TYPE "DT_PAR_PID_CROSS_FLOW_VALVE_1"
VERSION : 0.1
   STRUCT
      INPUT_RAMP_MIN_VAL { S7_SetPoint := 'False'} : "DT_PARAM_SOLO" := (FALSE, 832, 0, 0.0, 0, T#0MS, 0.0, 0.0, '%');
      INPUT_RAMP_MAX_VAL { S7_SetPoint := 'False'} : "DT_PARAM_SOLO" := (FALSE, 833, 0, 0.0, 0, T#0MS, 0.0, 0.0, '%');
      INPUT_RAMP_FALLING_TIME { S7_SetPoint := 'False'} : "DT_PARAM_SOLO" := (FALSE, 834, 0, 0.0, 0, T#0MS, 0.0, 0.0, 's');
      INPUT_RAMP_RISING_TIME { S7_SetPoint := 'False'} : "DT_PARAM_SOLO" := (FALSE, 835, 0, 0.0, 0, T#0MS, 0.0, 0.0, 's');
      OUTPUT_RAMP_FALLING_TIME { S7_SetPoint := 'False'} : "DT_PARAM_SOLO" := (FALSE, 836, 0, 0.0, 0, T#0MS, 0.0, 0.0, 's');
      OUTPUT_RAMP_RISING_TIME { S7_SetPoint := 'False'} : "DT_PARAM_SOLO" := (FALSE, 837, 0, 0.0, 0, T#0MS, 0.0, 0.0, 's');
      MAN_ON { S7_SetPoint := 'False'} : "DT_PARAM_SOLO" := (FALSE, 838, 1, 0.0, 0, T#0MS, 0.0, 0.0, '-');
      P_SEL { S7_SetPoint := 'False'} : "DT_PARAM_SOLO" := (FALSE, 839, 1, 0.0, 0, T#0MS, 0.0, 0.0, '-');
      I_SEL { S7_SetPoint := 'False'} : "DT_PARAM_SOLO" := (FALSE, 840, 1, 0.0, 0, T#0MS, 0.0, 0.0, '-');
      INT_HOLD { S7_SetPoint := 'False'} : "DT_PARAM_SOLO" := (FALSE, 841, 1, 0.0, 0, T#0MS, 0.0, 0.0, '-');
      D_SEL { S7_SetPoint := 'False'} : "DT_PARAM_SOLO" := (FALSE, 842, 1, 0.0, 0, T#0MS, 0.0, 0.0, '-');
      NUM_OF_CYCLES { S7_SetPoint := 'False'} : "DT_PARAM_SOLO" := (FALSE, 843, 1, 0.0, 0, T#0MS, 0.0, 0.0, '-');
      GAIN { S7_SetPoint := 'False'} : "DT_PARAM_SOLO" := (FALSE, 844, 0, 0.0, 0, T#0MS, 0.0, 0.0, '');
      TI { S7_SetPoint := 'False'} : "DT_PARAM_SOLO" := (FALSE, 845, 1, 0.0, 0, T#0MS, 0.0, 0.0, '-');
      TD { S7_SetPoint := 'False'} : "DT_PARAM_SOLO" := (FALSE, 846, 1, 0.0, 0, T#0MS, 0.0, 0.0, '-');
      TM_LAG { S7_SetPoint := 'False'} : "DT_PARAM_SOLO" := (FALSE, 847, 1, 300.0, 0, T#0MS, 0.0, 0.0, '-');
      DEAD_W { S7_SetPoint := 'False'} : "DT_PARAM_SOLO" := (FALSE, 848, 0, 100.0, 0, T#0MS, 0.0, 0.0, '%');
      LMN_HLM { S7_SetPoint := 'False'} : "DT_PARAM_SOLO" := (FALSE, 849, 0, 30.0, 0, T#0MS, 0.0, 0.0, '%');
      LMN_LLM { S7_SetPoint := 'False'} : "DT_PARAM_SOLO" := (FALSE, 850, 0, 300.0, 0, T#0MS, 0.0, 0.0, '%');
      REF_MIN_VAL { S7_SetPoint := 'False'} : "DT_PARAM_SOLO" := (FALSE, 851, 0, 0.0, 0, T#0MS, 0.0, 0.0, '%');
      REF_MAX_VAL { S7_SetPoint := 'False'} : "DT_PARAM_SOLO" := (FALSE, 852, 0, 0.0, 0, T#0MS, 0.0, 0.0, '%');
      LMN_FAC { S7_SetPoint := 'False'} : "DT_PARAM_SOLO" := (FALSE, 853, 0, 0.0, 0, T#0MS, 0.0, 0.0, '-');
      LMN_OFFSET { S7_SetPoint := 'False'} : "DT_PARAM_SOLO" := (FALSE, 854, 0, 0.0, 0, T#0MS, 0.0, 0.0, '%');
      DISV { S7_SetPoint := 'False'} : "DT_PARAM_SOLO" := (FALSE, 855, 0, 0.0, 0, T#0MS, 0.0, 0.0, '-');
      MAN { S7_SetPoint := 'False'} : "DT_PARAM_SOLO" := (FALSE, 856, 0, 0.0, 0, T#0MS, 0.0, 0.0, '%');
      REFERENCE_CORRECTION { S7_SetPoint := 'False'} : "DT_PARAM_SOLO" := (FALSE, 857, 0, 0.0, 0, T#0MS, 0.0, 0.0, '-');
      OUT_CTRL_MODE { S7_SetPoint := 'False'} : "DT_PARAM_SOLO" := (FALSE, 858, 1, 0.0, 0, T#0MS, 0.0, 0.0, '-');
      SPARE_4 { S7_SetPoint := 'False'} : "DT_PARAM_SOLO" := (FALSE, 859, 0, 0.0, 0, T#0MS, 0.0, 0.0, '');
      SPARE_5 { S7_SetPoint := 'False'} : "DT_PARAM_SOLO" := (FALSE, 860, 0, 0.0, 0, T#0MS, 0.0, 0.0, '');
      SPARE_6 { S7_SetPoint := 'False'} : "DT_PARAM_SOLO" := (FALSE, 861, 0, 0.0, 0, T#0MS, 0.0, 0.0, '');
      SPARE_7 { S7_SetPoint := 'False'} : "DT_PARAM_SOLO" := (FALSE, 862, 0, 0.0, 0, T#0MS, 0.0, 0.0, '');
      SPARE_8 { S7_SetPoint := 'False'} : "DT_PARAM_SOLO" := (FALSE, 863, 0, 0.0, 0, T#0MS, 0.0, 0.0, '');
   END_STRUCT;

END_TYPE

